RESOURCE RES0 : EMB_RES_ECO
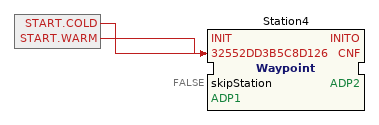
  FBS
    Station4 : Waypoint(skipStation := FALSE);
  END_FBS
  EVENT_CONNECTIONS
    START.COLD TO Station4.32552DD3B5C8D126;
    START.WARM TO Station4.32552DD3B5C8D126;
  END_CONNECTIONS
END_RESOURCE
